(* Schneider Machine Expert - Basic project Taimers_baise_and_signal_genarated, file version 2.9.0.0 *)
(* ProjectInformations: Name=New project *)

HARDWARE
  Cpu 0: TM221M16R/G
  EthernetConfiguration: NetworkName=M221, IpAllocationMode=FixedAddress, IpAddress=0.0.0.0, SubnetMask=0.0.0.0
  SerialLineConfiguration: Baud=Baud19200, Parity=ParityEven, DataBits=DataBits8, StopBits=StopBits1, PhysicalMedium=PhysicalMediumRs485, TransmissionMode=TransmissionModeModbusRtu, SlaveId=1, Addressing=SlaveAddressing
  MastTask: UsePeriodScanMode=false, PeriodScan=100
  FastTask: Period=255
  CpuBehavior: StartingMode=StartAsPreviousState, AutoSaveRamOnEeprom=true, WatchdogPeriod=250

SYMBOLS  (address, symbol, comment, settings)
  %M10      TON_START
  %M11      TON_OUT
  %M12      TOF_START
  %M13      TOF_OUT
  %M14      TON_START_SGD
  %M15      SET_UP_SIGNAL
  %M20      START_PID_GENERATED
  %TM0        [Type=TOF, Preset=50, Base=OneHundredMilliSeconds]
  %TM1        [Preset=50, Base=OneHundredMilliSeconds]
  %TM2        "SET_UP_SIGNAL_OFTER_1second"  [Preset=3, Base=OneSecond]
  %TM3        "SET_LOW_SIGNAL_ofter_one_second"  [Preset=3, Base=OneSecond]
  %TM4        "SET_UP_SIGN"  [Preset=3, Base=OneSecond]
  %TM5        "SET_LOW_SIGN"  [Type=TOF, Preset=3, Base=OneSecond]

POU New POU
  (* SectionNumber=1 *)

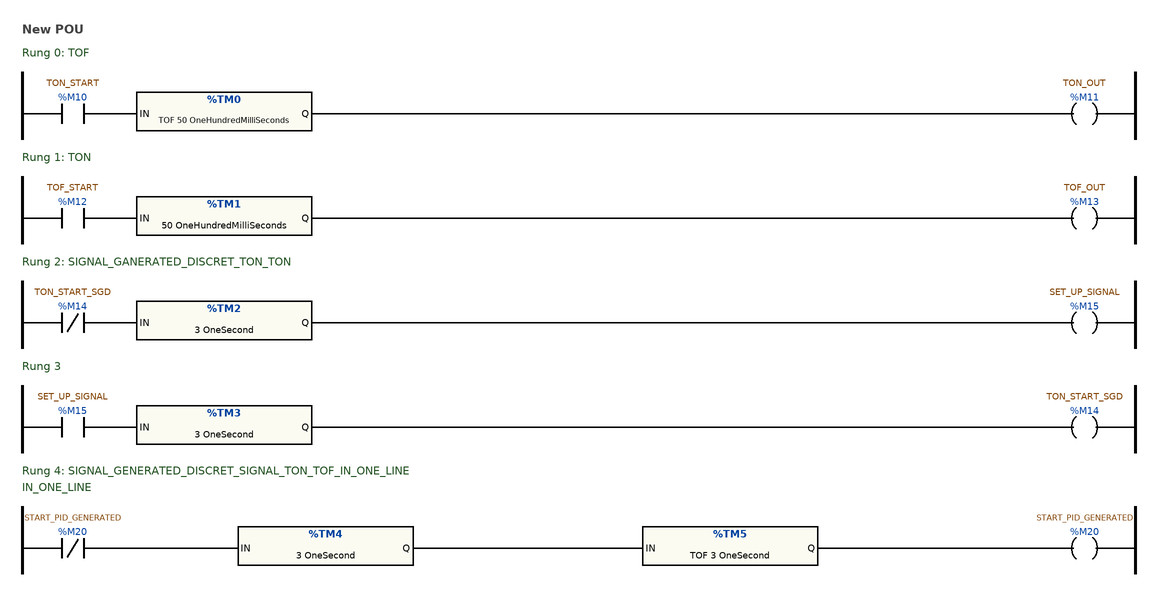

// Rung 0: TOF
  BLK %TM0
  LD %M10                 (* TON_START *)
  IN
  OUT_BLK
  LD Q
  ST %M11                 (* TON_OUT *)
  END_BLK
  // as ST:
  //   %TM0(IN := TON_START);
  //   TON_OUT := %TM0.Q;

// Rung 1: TON
  BLK %TM1
  LD %M12                 (* TOF_START *)
  IN
  OUT_BLK
  LD Q
  ST %M13                 (* TOF_OUT *)
  END_BLK
  // as ST:
  //   %TM1(IN := TOF_START);
  //   TOF_OUT := %TM1.Q;

// Rung 2: SIGNAL_GANERATED_DISCRET_TON_TON
  BLK %TM2
  LDN %M14                (* TON_START_SGD *)
  IN
  OUT_BLK
  LD Q
  ST %M15                 (* SET_UP_SIGNAL *)
  END_BLK
  // as ST:
  //   %TM2(IN := NOT TON_START_SGD);
  //   SET_UP_SIGNAL := %TM2.Q;

// Rung 3
  BLK %TM3
  LD %M15                 (* SET_UP_SIGNAL *)
  IN
  OUT_BLK
  LD Q
  ST %M14                 (* TON_START_SGD *)
  END_BLK
  // as ST:
  //   %TM3(IN := SET_UP_SIGNAL);
  //   TON_START_SGD := %TM3.Q;

// Rung 4: SIGNAL_GENERATED_DISCRET_SIGNAL_TON_TOF_IN_ONE_LINE
// IN_ONE_LINE
  LD 1
  MULTIFB
  BLK %TM4
  LD 1
  ANDN %M20               (* START_PID_GENERATED *)
  IN
  OUT_BLK
  LD Q
  ST %MW2009:X0
  END_BLK
  BLK %TM5
  LD %MW2009:X0
  IN
  OUT_BLK
  LD Q
  ST %M20                 (* START_PID_GENERATED *)
  END_BLK
  MULTIFB
  // as ST:
  //   %TM4(IN := NOT START_PID_GENERATED);
  //   %TM5(IN := %TM4.Q);
  //   START_PID_GENERATED := %TM5.Q;
